// TIA Portal V18 export
FUNCTION "VALIDACAO_ DOS_MODEZONES_ETR" : Void   // FC11, LAD
{ S7_Optimized_Access := 'TRUE' }
// stored: SetENOAutomatically false
   VAR_TEMP
      TESTE_1 : Bool;
      INDEX_STATION : Int;
      INDEX_POSITION : Int;
      INDEX_EQUIPMENT : Int;
      INDEX_SIGNAL : Int;
      leandro : Bool;
      index_positon_md1 : Int;
      index_equipament_md1 : Int;
      index_sinal_md1 : Int;
      POP_ID : String;
      BORDA : Bool;
      INDEX_CLEAN : Int;
      INDEX_FILA : Int;
      BORDA_1 : Bool;
      INDEX_SIGNAL1 : Int;
      INDEX_SIGNAL2 : Int;
      INDEX_VERIFICA : Int;
      barreira_invadida : Bool;
      aciona_buzzer : Bool;
      aciona_lampada_vermelha : Bool;
      aciona_lampada_verde : Bool;
      INTERLOCKS_MD1 : Bool;
      STATION : Int;
      SIGNAL : Int;
      EQUIPMENT : Int;
      count_LD : Bool;
      count_LE : Bool;
   END_VAR
   VAR_TEMP   // added for the SCL form of the ladder/FBD networks
      _w1 : Bool;
      _w2 : Bool;
   END_VAR
BEGIN

REGION Network 1: Buzzer
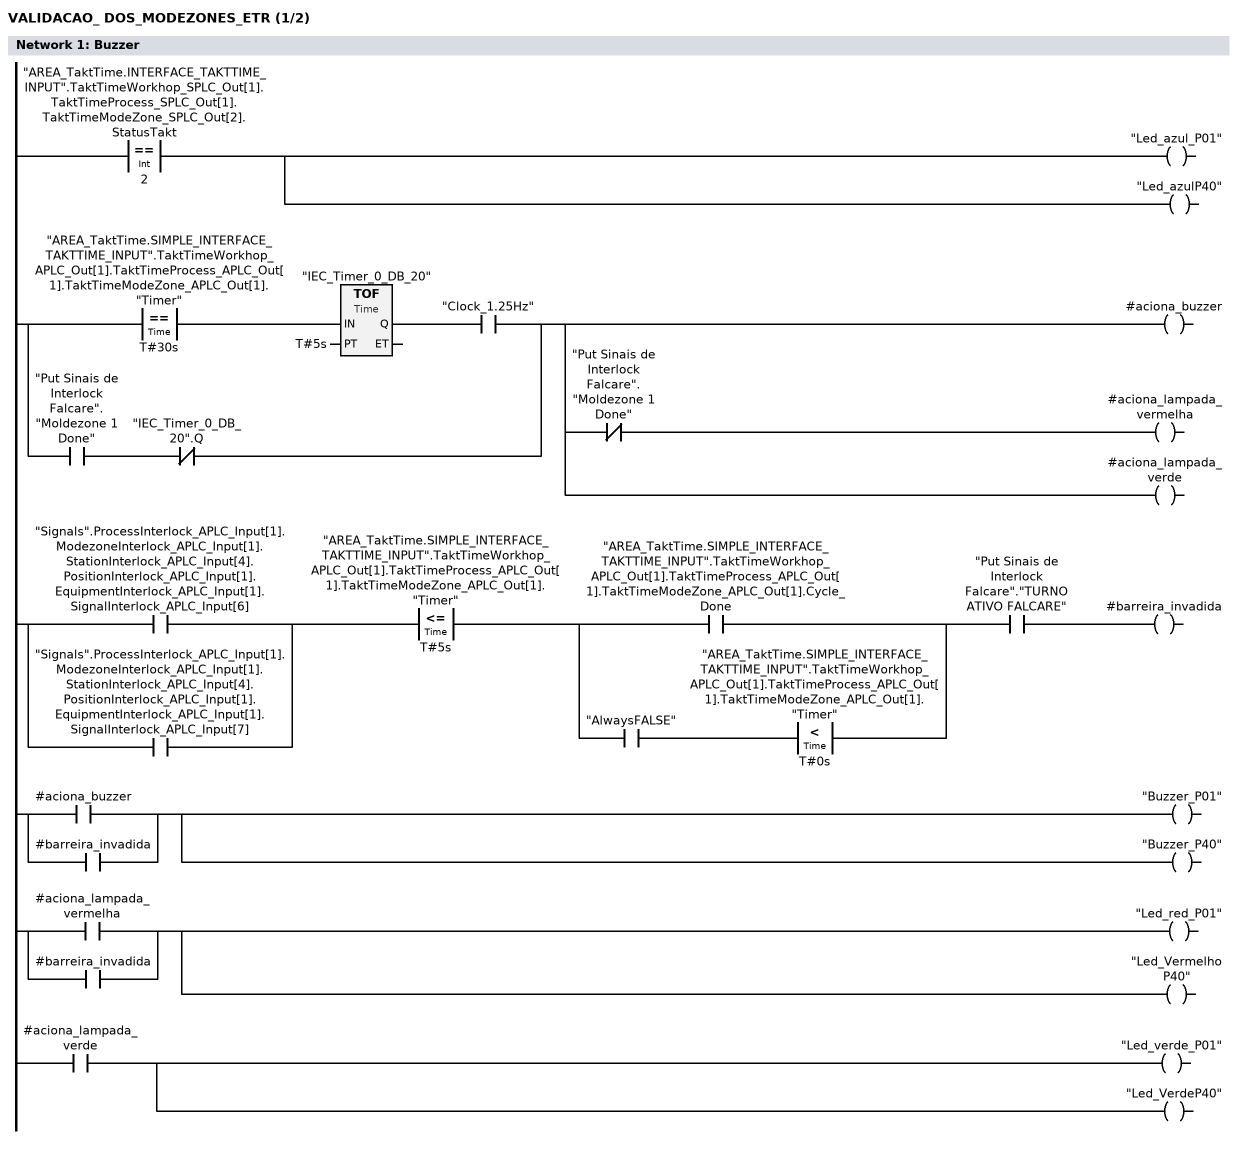
   RUNG wire#powerrail
      { S7_Templates := "SrcType := Int" } EQ_Contact(in1 := "AREA_TaktTime.INTERFACE_TAKTTIME_INPUT".TaktTimeWorkhop_SPLC_Out[1].TaktTimeProcess_SPLC_Out[1].TaktTimeModeZone_SPLC_Out[2].StatusTakt, in2 := 2)
      wire#w1
      Coil( "Led_azul_P01" )
   END_RUNG
   RUNG wire#w1
      Coil( "Led_azulP40" )
   END_RUNG
   RUNG wire#powerrail
      { S7_Templates := "SrcType := Time" } EQ_Contact(in1 := "AREA_TaktTime.SIMPLE_INTERFACE_TAKTTIME_INPUT".TaktTimeWorkhop_APLC_Out[1].TaktTimeProcess_APLC_Out[1].TaktTimeModeZone_APLC_Out[1]."Timer", in2 := T#30s)
      { S7_Templates := "time_type := Time" } "IEC_Timer_0_DB_20".TOF(pt := T#5s, et =>)
      Contact( "Clock_1.25Hz" )
      wire#w2
      Coil( #aciona_buzzer )
   END_RUNG
   RUNG wire#powerrail
      Contact( "Put Sinais de Interlock Falcare"."Moldezone 1 Done" )
      I_Contact( "IEC_Timer_0_DB_20".Q )
   END_RUNG wire#w2
   RUNG wire#w2
      I_Contact( "Put Sinais de Interlock Falcare"."Moldezone 1 Done" )
      Coil( #aciona_lampada_vermelha )
   END_RUNG
   RUNG wire#w2
      Coil( #aciona_lampada_verde )
   END_RUNG
   RUNG wire#powerrail
      Contact( "Signals".ProcessInterlock_APLC_Input[1].ModezoneInterlock_APLC_Input[1].StationInterlock_APLC_Input[4].PositionInterlock_APLC_Input[1].EquipmentInterlock_APLC_Input[1].SignalInterlock_APLC_Input[6] )
      wire#w3
      { S7_Templates := "SrcType := Time" } LE_Contact(in1 := "AREA_TaktTime.SIMPLE_INTERFACE_TAKTTIME_INPUT".TaktTimeWorkhop_APLC_Out[1].TaktTimeProcess_APLC_Out[1].TaktTimeModeZone_APLC_Out[1]."Timer", in2 := T#5s)
      wire#w4
      Contact( "AREA_TaktTime.SIMPLE_INTERFACE_TAKTTIME_INPUT".TaktTimeWorkhop_APLC_Out[1].TaktTimeProcess_APLC_Out[1].TaktTimeModeZone_APLC_Out[1].Cycle_Done )
      wire#w5
      Contact( "Put Sinais de Interlock Falcare"."TURNO ATIVO FALCARE" )
      Coil( #barreira_invadida )
   END_RUNG
   RUNG wire#powerrail
      Contact( "Signals".ProcessInterlock_APLC_Input[1].ModezoneInterlock_APLC_Input[1].StationInterlock_APLC_Input[4].PositionInterlock_APLC_Input[1].EquipmentInterlock_APLC_Input[1].SignalInterlock_APLC_Input[7] )
   END_RUNG wire#w3
   RUNG wire#w4
      Contact( "AlwaysFALSE" )
      { S7_Templates := "SrcType := Time" } LT_Contact(in1 := "AREA_TaktTime.SIMPLE_INTERFACE_TAKTTIME_INPUT".TaktTimeWorkhop_APLC_Out[1].TaktTimeProcess_APLC_Out[1].TaktTimeModeZone_APLC_Out[1]."Timer", in2 := T#0s)
   END_RUNG wire#w5
   RUNG wire#powerrail
      Contact( #aciona_buzzer )
      wire#w6
      Coil( "Buzzer_P01" )
   END_RUNG
   RUNG wire#powerrail
      Contact( #barreira_invadida )
   END_RUNG wire#w6
   RUNG wire#w6
      Coil( "Buzzer_P40" )
   END_RUNG
   RUNG wire#powerrail
      Contact( #aciona_lampada_vermelha )
      wire#w7
      Coil( "Led_red_P01" )
   END_RUNG
   RUNG wire#powerrail
      Contact( #barreira_invadida )
   END_RUNG wire#w7
   RUNG wire#w7
      Coil( "Led_VermelhoP40" )
   END_RUNG
   RUNG wire#powerrail
      Contact( #aciona_lampada_verde )
      wire#w8
      Coil( "Led_verde_P01" )
   END_RUNG
   RUNG wire#w8
      Coil( "Led_VerdeP40" )
   END_RUNG
   // the same network as SCL:
   "Led_azul_P01" := "AREA_TaktTime.INTERFACE_TAKTTIME_INPUT".TaktTimeWorkhop_SPLC_Out[1].TaktTimeProcess_SPLC_Out[1].TaktTimeModeZone_SPLC_Out[2].StatusTakt = 2;
   "Led_azulP40" := "Led_azul_P01";
   "IEC_Timer_0_DB_20".TOF(IN := "AREA_TaktTime.SIMPLE_INTERFACE_TAKTTIME_INPUT".TaktTimeWorkhop_APLC_Out[1].TaktTimeProcess_APLC_Out[1].TaktTimeModeZone_APLC_Out[1]."Timer" = T#30s,
                           PT := T#5s);
   #aciona_buzzer := ("IEC_Timer_0_DB_20".Q AND "Clock_1.25Hz") OR ("Put Sinais de Interlock Falcare"."Moldezone 1 Done" AND NOT "IEC_Timer_0_DB_20".Q);
   #aciona_lampada_vermelha := #aciona_buzzer AND NOT "Put Sinais de Interlock Falcare"."Moldezone 1 Done";
   #aciona_lampada_verde := #aciona_buzzer;
   #barreira_invadida := ("Signals".ProcessInterlock_APLC_Input[1].ModezoneInterlock_APLC_Input[1].StationInterlock_APLC_Input[4].PositionInterlock_APLC_Input[1].EquipmentInterlock_APLC_Input[1].SignalInterlock_APLC_Input[6] OR "Signals".ProcessInterlock_APLC_Input[1].ModezoneInterlock_APLC_Input[1].StationInterlock_APLC_Input[4].PositionInterlock_APLC_Input[1].EquipmentInterlock_APLC_Input[1].SignalInterlock_APLC_Input[7]) AND ("AREA_TaktTime.SIMPLE_INTERFACE_TAKTTIME_INPUT".TaktTimeWorkhop_APLC_Out[1].TaktTimeProcess_APLC_Out[1].TaktTimeModeZone_APLC_Out[1]."Timer" <= T#5s) AND ("AREA_TaktTime.SIMPLE_INTERFACE_TAKTTIME_INPUT".TaktTimeWorkhop_APLC_Out[1].TaktTimeProcess_APLC_Out[1].TaktTimeModeZone_APLC_Out[1].Cycle_Done OR ("AlwaysFALSE" AND ("AREA_TaktTime.SIMPLE_INTERFACE_TAKTTIME_INPUT".TaktTimeWorkhop_APLC_Out[1].TaktTimeProcess_APLC_Out[1].TaktTimeModeZone_APLC_Out[1]."Timer" < T#0s))) AND "Put Sinais de Interlock Falcare"."TURNO ATIVO FALCARE";
   "Buzzer_P01" := #aciona_buzzer OR #barreira_invadida;
   "Buzzer_P40" := "Buzzer_P01";
   "Led_red_P01" := #aciona_lampada_vermelha OR #barreira_invadida;
   "Led_VermelhoP40" := "Led_red_P01";
   "Led_verde_P01" := #aciona_lampada_verde;
   "Led_VerdeP40" := #aciona_lampada_verde;
END_REGION

REGION Network 2 (SCL)
   IF "VERIFICA INTERLOCK"."ATIVA FOR" THEN
       FOR #INDEX_SIGNAL := 1 TO "Station_Setup_Const" DO
           FOR #INDEX_SIGNAL1 := 1 TO "Equipment_Setup_Const" DO
               FOR #INDEX_SIGNAL2 := 1 TO "Signal_Setup_Const" DO
                   IF "Signals".ProcessInterlock_APLC_Input[1].ModezoneInterlock_APLC_Input[2].StationInterlock_APLC_Input[#INDEX_SIGNAL]
                       .PositionInterlock_APLC_Input[1].EquipmentInterlock_APLC_Input[#INDEX_SIGNAL1].SignalInterlock_APLC_Input[#INDEX_SIGNAL2] = TRUE THEN
                       FOR #INDEX_VERIFICA := 1 TO 10 DO
                           IF "VERIFICA INTERLOCK".INTERLOCK[#INDEX_VERIFICA].STATION = 0 THEN
                               "VERIFICA INTERLOCK".INTERLOCK[#INDEX_VERIFICA].STATION := #INDEX_SIGNAL;
                               "VERIFICA INTERLOCK".INTERLOCK[#INDEX_VERIFICA].EQUIPAMENTO := #INDEX_SIGNAL1;
                               "VERIFICA INTERLOCK".INTERLOCK[#INDEX_VERIFICA].SINAL := #INDEX_SIGNAL2;
                               EXIT;
                           END_IF;
                       END_FOR;
                   END_IF;
                   END_FOR;
               END_FOR;
           END_FOR;
           "VERIFICA INTERLOCK"."ATIVA FOR" := FALSE;
       END_IF;
END_REGION

REGION Network 3
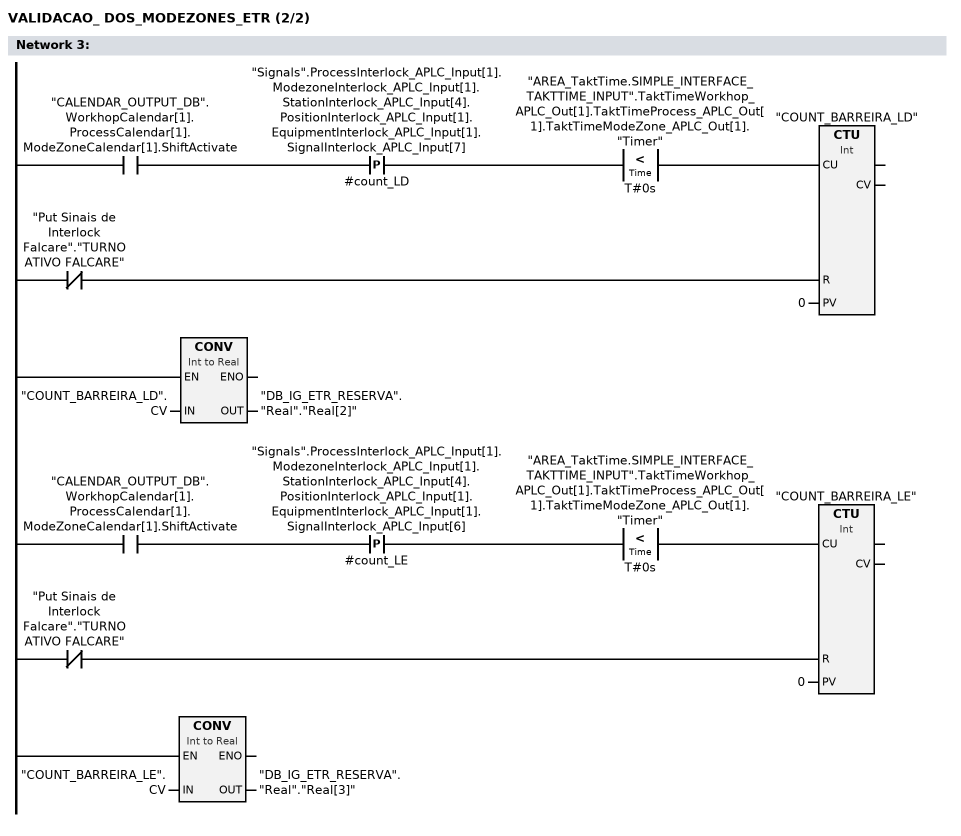
   RUNG wire#powerrail
      Contact( "CALENDAR_OUTPUT_DB".WorkhopCalendar[1].ProcessCalendar[1].ModeZoneCalendar[1].ShiftActivate )
      P_Contact(operand := "Signals".ProcessInterlock_APLC_Input[1].ModezoneInterlock_APLC_Input[1].StationInterlock_APLC_Input[4].PositionInterlock_APLC_Input[1].EquipmentInterlock_APLC_Input[1].SignalInterlock_APLC_Input[7], bit := #count_LD)
      { S7_Templates := "SrcType := Time" } LT_Contact(in1 := "AREA_TaktTime.SIMPLE_INTERFACE_TAKTTIME_INPUT".TaktTimeWorkhop_APLC_Out[1].TaktTimeProcess_APLC_Out[1].TaktTimeModeZone_APLC_Out[1]."Timer", in2 := T#0s)
      { S7_Templates := "value_type := Int" } "COUNT_BARREIRA_LD".CTU(r := wire#w1, pv := 0, cv =>)
   END_RUNG
   RUNG wire#powerrail
      I_Contact( "Put Sinais de Interlock Falcare"."TURNO ATIVO FALCARE" )
   END_RUNG wire#w1
   RUNG wire#powerrail
      { S7_Templates := "[SrcType := Int, DestType := Real]" } Convert(in := "COUNT_BARREIRA_LD".CV, out => "DB_IG_ETR_RESERVA"."Real"."Real[2]")
   END_RUNG
   RUNG wire#powerrail
      Contact( "CALENDAR_OUTPUT_DB".WorkhopCalendar[1].ProcessCalendar[1].ModeZoneCalendar[1].ShiftActivate )
      P_Contact(operand := "Signals".ProcessInterlock_APLC_Input[1].ModezoneInterlock_APLC_Input[1].StationInterlock_APLC_Input[4].PositionInterlock_APLC_Input[1].EquipmentInterlock_APLC_Input[1].SignalInterlock_APLC_Input[6], bit := #count_LE)
      { S7_Templates := "SrcType := Time" } LT_Contact(in1 := "AREA_TaktTime.SIMPLE_INTERFACE_TAKTTIME_INPUT".TaktTimeWorkhop_APLC_Out[1].TaktTimeProcess_APLC_Out[1].TaktTimeModeZone_APLC_Out[1]."Timer", in2 := T#0s)
      { S7_Templates := "value_type := Int" } "COUNT_BARREIRA_LE".CTU(r := wire#w2, pv := 0, cv =>)
   END_RUNG
   RUNG wire#powerrail
      I_Contact( "Put Sinais de Interlock Falcare"."TURNO ATIVO FALCARE" )
   END_RUNG wire#w2
   RUNG wire#powerrail
      { S7_Templates := "[SrcType := Int, DestType := Real]" } Convert(in := "COUNT_BARREIRA_LE".CV, out => "DB_IG_ETR_RESERVA"."Real"."Real[3]")
   END_RUNG
   // the same network as SCL:
   #_w1 := "CALENDAR_OUTPUT_DB".WorkhopCalendar[1].ProcessCalendar[1].ModeZoneCalendar[1].ShiftActivate AND "Signals".ProcessInterlock_APLC_Input[1].ModezoneInterlock_APLC_Input[1].StationInterlock_APLC_Input[4].PositionInterlock_APLC_Input[1].EquipmentInterlock_APLC_Input[1].SignalInterlock_APLC_Input[7] AND NOT #count_LD;   // rising edge of "Signals".ProcessInterlock_APLC_Input[1].ModezoneInterlock_APLC_Input[1].StationInterlock_APLC_Input[4].PositionInterlock_APLC_Input[1].EquipmentInterlock_APLC_Input[1].SignalInterlock_APLC_Input[7]
   #count_LD := "Signals".ProcessInterlock_APLC_Input[1].ModezoneInterlock_APLC_Input[1].StationInterlock_APLC_Input[4].PositionInterlock_APLC_Input[1].EquipmentInterlock_APLC_Input[1].SignalInterlock_APLC_Input[7];
   "COUNT_BARREIRA_LD".CTU(CU := #_w1 AND ("AREA_TaktTime.SIMPLE_INTERFACE_TAKTTIME_INPUT".TaktTimeWorkhop_APLC_Out[1].TaktTimeProcess_APLC_Out[1].TaktTimeModeZone_APLC_Out[1]."Timer" < T#0s),
                           R := NOT "Put Sinais de Interlock Falcare"."TURNO ATIVO FALCARE",
                           PV := 0);
   "DB_IG_ETR_RESERVA"."Real"."Real[2]" := INT_TO_REAL("COUNT_BARREIRA_LD".CV);
   #_w2 := "CALENDAR_OUTPUT_DB".WorkhopCalendar[1].ProcessCalendar[1].ModeZoneCalendar[1].ShiftActivate AND "Signals".ProcessInterlock_APLC_Input[1].ModezoneInterlock_APLC_Input[1].StationInterlock_APLC_Input[4].PositionInterlock_APLC_Input[1].EquipmentInterlock_APLC_Input[1].SignalInterlock_APLC_Input[6] AND NOT #count_LE;   // rising edge of "Signals".ProcessInterlock_APLC_Input[1].ModezoneInterlock_APLC_Input[1].StationInterlock_APLC_Input[4].PositionInterlock_APLC_Input[1].EquipmentInterlock_APLC_Input[1].SignalInterlock_APLC_Input[6]
   #count_LE := "Signals".ProcessInterlock_APLC_Input[1].ModezoneInterlock_APLC_Input[1].StationInterlock_APLC_Input[4].PositionInterlock_APLC_Input[1].EquipmentInterlock_APLC_Input[1].SignalInterlock_APLC_Input[6];
   "COUNT_BARREIRA_LE".CTU(CU := #_w2 AND ("AREA_TaktTime.SIMPLE_INTERFACE_TAKTTIME_INPUT".TaktTimeWorkhop_APLC_Out[1].TaktTimeProcess_APLC_Out[1].TaktTimeModeZone_APLC_Out[1]."Timer" < T#0s),
                           R := NOT "Put Sinais de Interlock Falcare"."TURNO ATIVO FALCARE",
                           PV := 0);
   "DB_IG_ETR_RESERVA"."Real"."Real[3]" := INT_TO_REAL("COUNT_BARREIRA_LE".CV);
END_REGION
END_FUNCTION
